(* IEC 61131-3 sources: 2026_Projet_YGO_ExcavatriceDragage/TOOLS/TEST_AUTO_CI/RESULTS/_TROUBLESHOOTING/AGY02_T417_M3_SANDBOX, 1 file *)

(* ---- test_m3_sandbox.st ---- *)
SETUP
VAR
    FB : FB_TestHarnessT417_M3;
    RawPosM1 : UDINT := 0;
    RawPosM2 : UDINT := 0;
END_VAR
END_SETUP

TEST 'SANDBOX-M3-01 Approche Manu vers Tremie (baseline simu)'
VAR
    i : INT;
END_VAR
    FOR i := 1 TO 320 DO
        ADVANCE_TIME(10000000);
        FB(Enable := TRUE, StepForceTgt := -1, SimM3Slope_Mps2 := 0.0, BenneDone := FALSE, BenneIsOpen := FALSE);
    END_FOR;
    ASSERT_NEAR(FB.M3PositionTrue_M, 5.0, 0.05, 'Depart P1');

    (* Deplacement vers Tremie en Manu (JoystickLeft) : 5.0 m a 0.20 m/s -> ~25 s *)
    FOR i := 1 TO 3000 DO
        ADVANCE_TIME(10000000);
        FB(Enable := TRUE, StepForceTgt := -1, JoystickLeft := TRUE, SimM3Slope_Mps2 := 0.0, BenneDone := FALSE, BenneIsOpen := FALSE);
    END_FOR;
    ASSERT_TRUE(FB.M3AtTremie, 'Capteur Tremie atteint');
    ASSERT_GT(FB.M3PositionTrue_M, -0.45, 'Simu actuelle s arrete avant la butee mecanique -0.50m');
END_TEST
